Fanuc KAREL source: kt00883.KL

-- PROVISIONAL review KL for V940-1; original PC SHA256 10e974c0ff72d3aa6bd7739ad74bb5f92644f4e6e3ec01b2cfe82fdf2f614aae
-- Incomplete behavior may be omitted. Consult companion uncertainty JSON. Do not deploy.
PROGRAM KT00883
%NOLOCKGROUP
VAR
  R1 : REAL
  R2 : REAL
  OUT : REAL
BEGIN
  -- V9_ZERO_TABLE_METADATA_HINT layout=0001; no indexed target words; source/name/runtime held
  -- UNRESOLVED_PC offsets 5-16; opcodes 2E,23
  -- UNRESOLVED_PC offsets 21-32; opcodes 2E,23
  -- UNRESOLVED_PC offsets 37-48; opcodes 2E,23
  -- UNRESOLVED_PC offsets 53-64; opcodes 2E,23
  -- UNRESOLVED_PC offsets 69-90; opcodes 27,22,22,76,23
  -- UNRESOLVED_PC offsets 95-99; opcodes 7F
END KT00883
